(* Logix 5000 project; controller lab_5 vendor 1 type 14 code 149 rev 32.11; software revision 32.00 *)

TASK MainTask (continuous, watchdog 500 ms) : MainProgram

MODULES
   Local : vendor 1 type 14 code 149 (Compact 0, rev 32.11)
      Discrete_IO : Embedded (Compact 1, rev 3.1, Output RPI 20 ms)
END_MODULES

PROGRAM MainProgram   (* main routine MainRoutine *)
VAR
   e_stop : ALIAS FOR Local:1:I.Data.0;
   green_light : ALIAS FOR Local:1:O.Data.2;
   motor : ALIAS FOR Local:1:O.Data.6;
   red_light : ALIAS FOR Local:1:O.Data.0;
   start_button : ALIAS FOR Local:1:I.Data.2;
   stop_button : ALIAS FOR Local:1:I.Data.1;
   system_run : BOOL;
   timer : TIMER := (PRE := 5000);
END_VAR

ROUTINE MainRoutine   (* ladder *)
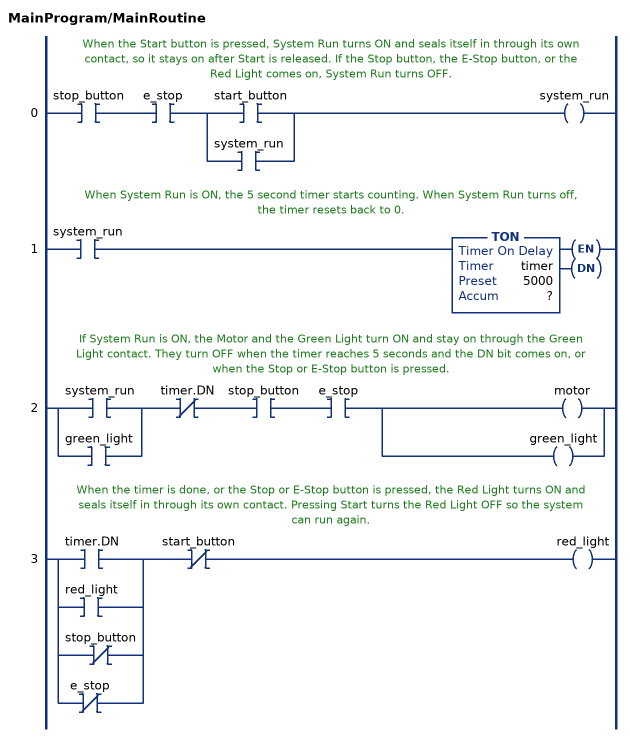
   // When the Start button is pressed, System Run turns ON and seals itself in through its own contact, so it stays on after Start is released. If the Stop button, the E-Stop button, or the Red Light comes on, System Run turns OFF.
   0: XIC(stop_button)XIC(e_stop)[XIC(start_button) ,XIC(system_run) ]OTE(system_run);
   // When System Run is ON, the 5 second timer starts counting. When System Run turns off, the timer resets back to 0.
   1: XIC(system_run)TON(timer,?,?);
   // If System Run is ON, the Motor and the Green Light turn ON and stay on through the Green Light contact. They turn OFF when the timer reaches 5 seconds and the DN bit comes on, or when the Stop or E-Stop button is pressed.
   2: [XIC(system_run) ,XIC(green_light) ]XIO(timer.DN)XIC(stop_button)XIC(e_stop)[OTE(motor) ,OTE(green_light) ];
   // When the timer is done, or the Stop or E-Stop button is pressed, the Red Light turns ON and seals itself in through its own contact. Pressing Start turns the Red Light OFF so the system can run again.
   3: [[[XIC(timer.DN) ,XIC(red_light) ] ,XIO(stop_button) ] ,XIO(e_stop) ]XIO(start_button)OTE(red_light);
END_ROUTINE
END_PROGRAM
